PROGRAM main
  VAR
    S1 AT %IX0.0  : BOOL; (* abrir, NA *)
    S2 AT %IX0.1  : BOOL; (* cerrar, NA *)
    S0 AT %IX0.2  : BOOL; (* parada, NC: TRUE sin pulsar *)
    B1 AT %IX0.3  : BOOL; (* final: portón abierto *)
    B2 AT %IX0.4  : BOOL; (* final: portón cerrado *)
    B3 AT %IX0.5  : BOOL; (* barrera: obstáculo en el paso *)
    KM1 AT %QX0.0 : BOOL; (* motor: abrir *)
    KM2 AT %QX0.1 : BOOL; (* motor: cerrar *)
    H1 AT %QX0.2  : BOOL; (* baliza de movimiento *)
    ETAPA         : INT; (* 0 parado, 1 abriendo, 2 cerrando *)
    E0            : BOOL; (* ETAPA = 0 *)
    E1            : BOOL; (* ETAPA = 1 *)
    E2            : BOOL; (* ETAPA = 2 *)
  END_VAR

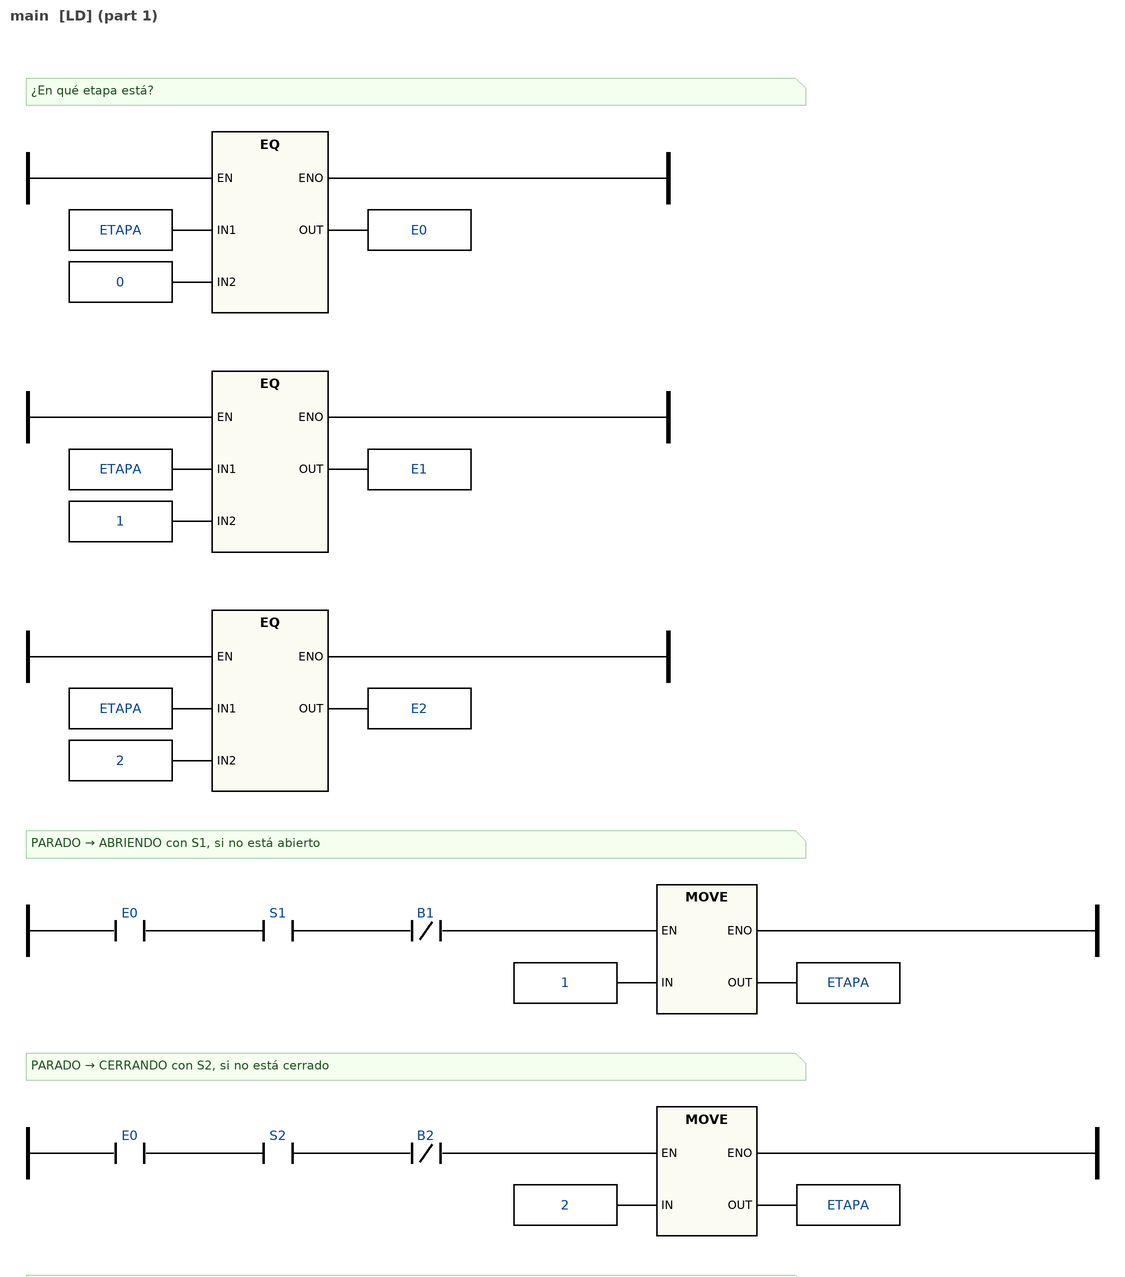
(* LD diagram, written out as Structured Text *)
(* ¿En qué etapa está? *)
E0 := ETAPA = 0;
E1 := ETAPA = 1;
E2 := ETAPA = 2;
(* PARADO → ABRIENDO con S1, si no está abierto *)
IF E0 AND S1 AND NOT B1 THEN ETAPA := 1; END_IF;
(* PARADO → CERRANDO con S2, si no está cerrado *)
IF E0 AND S2 AND NOT B2 THEN ETAPA := 2; END_IF;
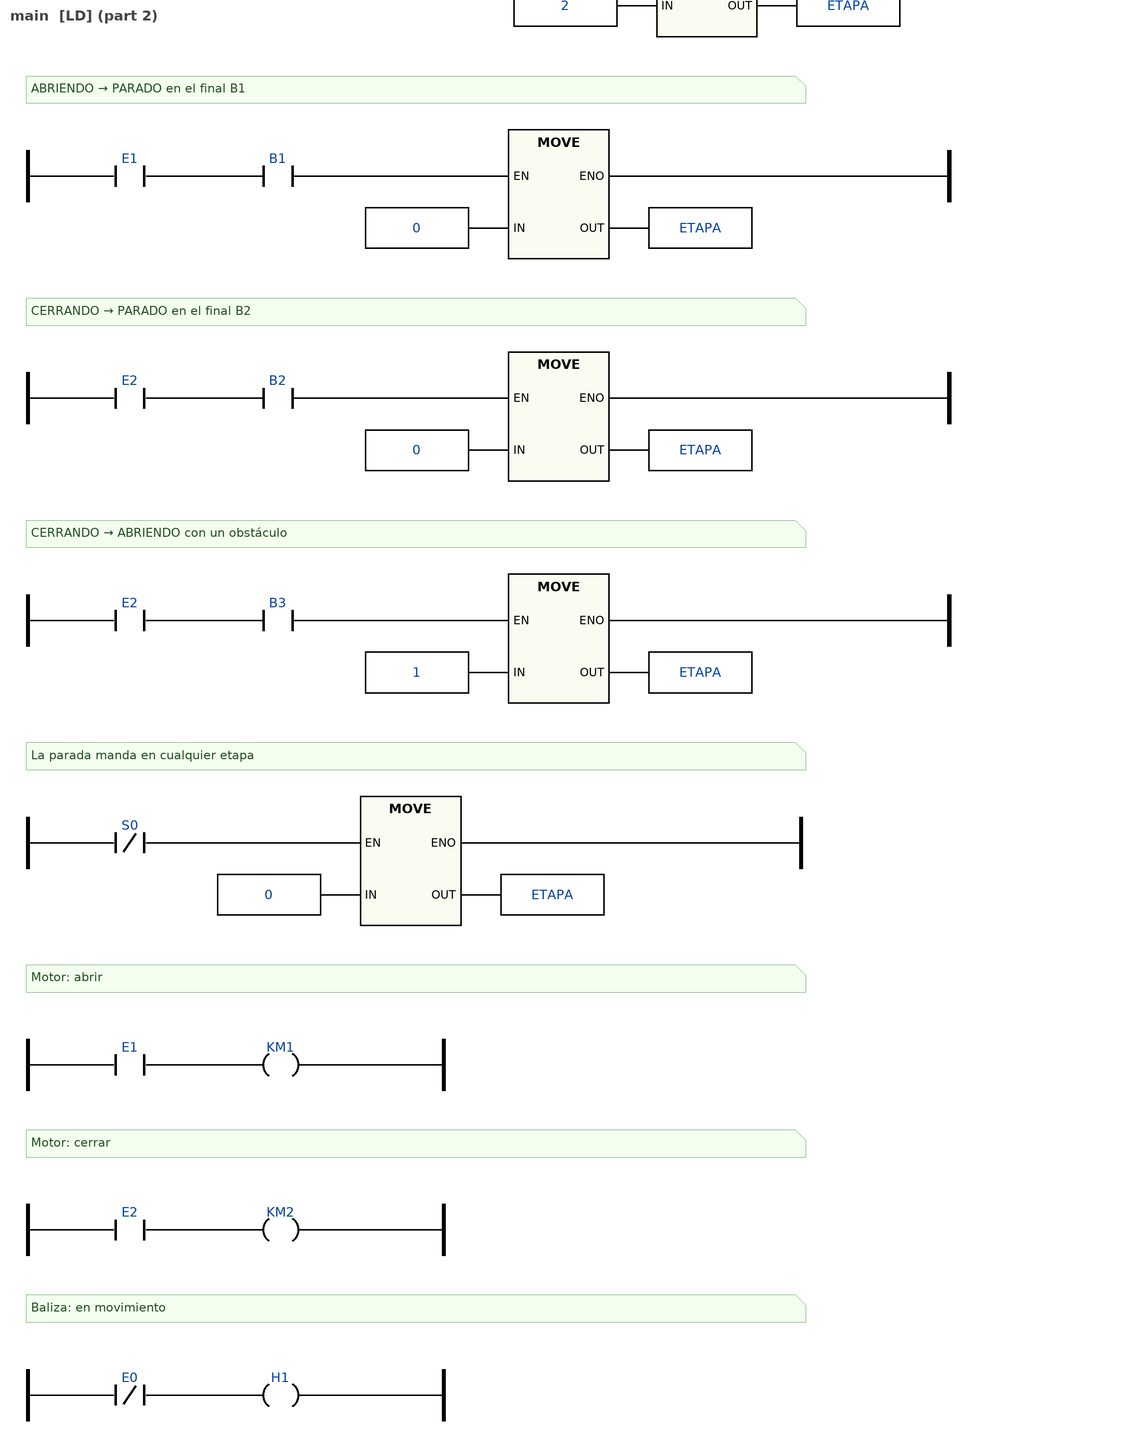
(* ABRIENDO → PARADO en el final B1 *)
IF E1 AND B1 THEN ETAPA := 0; END_IF;
(* CERRANDO → PARADO en el final B2 *)
IF E2 AND B2 THEN ETAPA := 0; END_IF;
(* CERRANDO → ABRIENDO con un obstáculo *)
IF E2 AND B3 THEN ETAPA := 1; END_IF;
(* La parada manda en cualquier etapa *)
IF NOT S0 THEN ETAPA := 0; END_IF;
(* Motor: abrir *)
KM1 := E1;
(* Motor: cerrar *)
KM2 := E2;
(* Baliza: en movimiento *)
H1 := NOT E0;
END_PROGRAM
